Staubli VAL3: utEvents.dtx

public bool bClick
public bool bMouseDown
public bool bMouseUp
